FUNCTION_BLOCK fbBistableSingleCoilRelay IMPLEMENTS iRelay
VAR
	RelayOutput AT %Q* : BOOL;

    PulseReq : BOOL;
    PulseTP : TP;
	
	ToggleVirtualStateTrig : R_TRIG;
END_VAR
VAR CONSTANT
    PulseTime : TIME := T#200MS;
END_VAR
VAR PERSISTENT
	RelaySet : BOOL;
END_VAR

(* 
	NOTE:
	After power reset, state of the relay is unknown and RelaySet variable may keep wrong value. 
	If RelaySet doesn't reflect the actual, physical state of relay, methods Reset() and Set() will have reverse effect.
	
	POSSIBLE SOLUTIONS:
	- relay state feedback as physical input signal
	- additional variable/method to toggle RelaySet without changing physical output RelayOutput
		implemented ToggleVirtualState(Execute : BOOL)
*)

PulseTP(IN := PulseReq, PT := PulseTime);
RelayOutput := PulseTP.Q;

IF PulseReq THEN
	RelaySet := NOT RelaySet;
	PulseReq := FALSE;
END_IF

{warning 'Add property implementation'}
PROPERTY IsSet : BOOL
GET
IsSet := RelaySet;
END_GET
END_PROPERTY

{warning 'Add method implementation '}
METHOD Reset
IF RelaySet THEN
	PulseReq := TRUE;	
END_IF
END_METHOD

{warning 'Add method implementation '}
METHOD Set
IF NOT RelaySet THEN
	PulseReq := TRUE;	
END_IF
END_METHOD

METHOD ToggleVirtualState
VAR_INPUT
    Execute : BOOL;
END_VAR
(*
	Do not call it conditionally ( inside IF )
	Works best when called every PLC cycle
*)


ToggleVirtualStateTrig(CLK := Execute);
IF ToggleVirtualStateTrig.Q THEN
	THIS^.RelaySet := NOT THIS^.RelaySet;
END_IF
END_METHOD

END_FUNCTION_BLOCK

(* stored: Version 1.1.0.1
   POU fbBistableSingleCoilRelay: Id {0fae3c70-2fb9-46ef-aed9-dd8518f75f14}, SpecialFunc None
   Property IsSet: Id {6eb00f3d-c6aa-447e-be14-295ed0b97da3}
   Get Get: Id {8141aa7c-5d5a-4692-8792-e740038cfeb1}
   Method Reset: Id {a9ee56df-9b3e-4fd0-adec-58152da57428}
   Method Set: Id {e2e6b3f1-b1b7-4ef5-8c82-af292b3e5831}
   Method ToggleVirtualState: Id {fce4026f-45b5-4475-b209-29bf29b1bc0f} *)
